// TIA Portal V21 export
Screen "T03_Btn"  1024x768, Number=23
  ScreenLayer 
    Button "P_Btn" at 0,0 size 100x30  TextOff="BTN", TextOn="BTN"
